Fanuc KAREL source: kt00186.KL

-- PROVISIONAL review KL for V940-1; original PC SHA256 a36a5d9d5ca2b54fecbe29b888652f7c3b1ce0d94afe67aa2a71675b8d8bd79f
-- Incomplete behavior may be omitted. Consult companion uncertainty JSON. Do not deploy.
PROGRAM KT00186
%NOLOCKGROUP
VAR
  I2 : INTEGER
  OUT : REAL
-- UNRESOLVED_DECL H1 type=002017
BEGIN
  -- V9_ZERO_TABLE_METADATA_HINT layout=0001; no indexed target words; source/name/runtime held
  -- UNRESOLVED_PC offsets 5-19; opcodes 2E,22,9D,33,B4
  -- UNRESOLVED_PC offsets 24-35; opcodes 2E,23
  -- UNRESOLVED_PC offsets 40-63; opcodes 22,9D,33,B3,21,56,64,23
  -- UNRESOLVED_PC offsets 68-72; opcodes 7F
END KT00186
